// TIA Portal project "Hardware" (V21)

(* hardware
DEVICE "Controller"  S7-1500 station
   slot 0: "Rail_0"  Rack  6ES7 590-1***0-0AA0
   slot 1: "Controller"  CPU 1516-3 PN/DP  6ES7 516-3AN02-0AB0  V2.9
      slot 3: "CPU display_1"  6ES7591-1BA00-0AA0
      slot 32768: "PROFINET interface_1"  X1
         slot 32769: "Port_1"  X1 P1
         slot 32770: "Port_2"  X1 P2
      slot 33024: "PROFINET interface_2"  X2
         slot 33025: "Port_1"  X2 P1
      slot 33280: "DP interface_1"  X3
      slot 34817: "Virtual CP interface port_1"  Virtual CP interface port  Virtual CP interface port
   slot 2: "DI_Main"  DI 32x24VDC HF  6ES7 521-1BL00-0AB0  V2.2
   slot 3: "DQ_Main"  DQ 32x24VDC/0.5A HF  6ES7 522-1BL01-0AB0  V1.1
   slot 4: "AI_Main"  AI 8xU/I/RTD/TC ST  6ES7 531-7KF00-0AB0  V2.2
   slot 5: "AQ_Main"  AQ 4xU/I ST  6ES7 532-5HD00-0AB0  V2.2
DEVICE "Remote_PN_1"  ET 200SP-Station
   slot 0: "Rack_0"  Rack  6ES5 710-8MAx1
   slot 0: "Remote_PN_1"  IM 155-6 PN ST  6ES7 155-6AU01-0BN0  V4.2
   slot 1: "Inputs_1"  DI 8x24VDC ST  6ES7 131-6BF01-0BA0  V0.0
      slot 1: "Inputs_1"  DI 8x24VDC ST
   slot 2: "Outputs_1"  DQ 8x24VDC/0.5A ST  6ES7 132-6BF01-0BA0  V0.0
      slot 1: "Outputs_1"  DQ 8x24VDC/0.5A ST
   slot 3: "Analog_1"  AI 4xI 2-,4-wire ST  6ES7 134-6GD01-0BA1  V2.0
      slot 1: "Analog_1"  AI 4xI 2-,4-wire ST
   slot 127: "BA 2xRJ45"  BA 2xRJ45  6ES7 193-6AR00-0AA0  V0.0
      slot 1: "Port_1"  X1 P1R  6ES7 193-6AR00-0AA0  V0.0
      slot 2: "Port_2"  X1 P2R  6ES7 193-6AR00-0AA0  V0.0
DEVICE "Remote_PN_2"  ET 200SP-Station
   slot 0: "Rack_0"  Rack  6ES5 710-8MAx1
   slot 0: "Remote_PN_2"  IM 155-6 PN ST  6ES7 155-6AU01-0BN0  V4.2
   slot 1: "Inputs_2"  DI 8x24VDC ST  6ES7 131-6BF01-0BA0  V0.0
      slot 1: "Inputs_2"  DI 8x24VDC ST
   slot 127: "BA 2xRJ45"  BA 2xRJ45  6ES7 193-6AR00-0AA0  V0.0
      slot 1: "Port_1"  X1 P1R  6ES7 193-6AR00-0AA0  V0.0
      slot 2: "Port_2"  X1 P2R  6ES7 193-6AR00-0AA0  V0.0
DEVICE "Remote_DP"  ET 200SP-Station
   slot 0: "Rack_0"  Rack  6ES5 710-8MAx1
   slot 0: "Remote_DP"  IM 155-6 DP HF  6ES7 155-6BU01-0CN0  V4.2
   slot 1: "Inputs_DP"  DI 8x24VDC ST  6ES7 131-6BF01-0BA0  V0.0
      slot 1: "Inputs_DP"  DI 8x24VDC ST
   slot 2: "Outputs_DP"  DQ 8x24VDC/0.5A ST  6ES7 132-6BF01-0BA0  V0.0
      slot 1: "Outputs_DP"  DQ 8x24VDC/0.5A ST
DEVICE "Partner"  S7-1500 station
   slot 0: "Rail_0"  Rack  6ES7 590-1***0-0AA0
   slot 1: "Partner"  CPU 1511-1 PN  6ES7 511-1AK02-0AB0  V2.9
      slot 3: "CPU display_1"  6ES7591-1AA00-0AA0
      slot 32768: "PROFINET interface_1"  X1
         slot 32769: "Port_1"  X1 P1
         slot 32770: "Port_2"  X1 P2
      slot 34817: "Virtual CP interface port_1"  Virtual CP interface port  Virtual CP interface port
DEVICE "Partner_IO"  ET 200SP-Station
   slot 0: "Rack_0"  Rack  6ES5 710-8MAx1
   slot 0: "Partner_IO"  IM 155-6 PN ST  6ES7 155-6AU01-0BN0  V4.2
   slot 1: "Outputs_P"  DQ 8x24VDC/0.5A ST  6ES7 132-6BF01-0BA0  V0.0
      slot 1: "Outputs_P"  DQ 8x24VDC/0.5A ST
   slot 127: "BA 2xRJ45"  BA 2xRJ45  6ES7 193-6AR00-0AA0  V0.0
      slot 1: "Port_1"  X1 P1R  6ES7 193-6AR00-0AA0  V0.0
      slot 2: "Port_2"  X1 P2R  6ES7 193-6AR00-0AA0  V0.0
DEVICE "Spare_PN"  ET 200SP-Station
   slot 0: "Rack_0"  Rack  6ES5 710-8MAx1
   slot 0: "Spare_PN"  IM 155-6 PN ST  6ES7 155-6AU01-0BN0  V4.2
   slot 1: "Inputs_S"  DI 8x24VDC ST  6ES7 131-6BF01-0BA0  V0.0
      slot 1: "Inputs_S"  DI 8x24VDC ST
   slot 127: "BA 2xRJ45"  BA 2xRJ45  6ES7 193-6AR00-0AA0  V0.0
      slot 1: "Port_1"  X1 P1R  6ES7 193-6AR00-0AA0  V0.0
      slot 2: "Port_2"  X1 P2R  6ES7 193-6AR00-0AA0  V0.0
*)

// ===== PLC "Controller"  CPU 1516-3 PN/DP =====

VAR_GLOBAL   // PLC tag table "IO"
   "Start_Line" AT %I10.0 : Bool;   // First input of DI_Main
   "Lamp_Line" AT %Q0.0 : Bool;   // First output of DQ_Main
END_VAR

ORGANIZATION_BLOCK "Main"   // OB1, SCL, ProgramCycle
TITLE = "Main Program Sweep (Cycle)"
{ S7_Optimized_Access := 'TRUE' }
VERSION : 0.1
   VAR_INPUT
      Initial_Call : Bool;   // Initial call of this OB
      Remanence : Bool;   // =True, if remanent data are available
   END_VAR
BEGIN

    "Lamp_Line" := "Start_Line";
END_ORGANIZATION_BLOCK

// ===== PLC "Partner"  CPU 1511-1 PN =====

VAR_GLOBAL   // PLC tag table "IO"
   "Start_Partner" AT %I0.0 : Bool;   // An input of the partner
   "Lamp_Partner" AT %Q0.0 : Bool;   // First output of Outputs_P
END_VAR

ORGANIZATION_BLOCK "Main"   // OB1, SCL, ProgramCycle
TITLE = "Main Program Sweep (Cycle)"
{ S7_Optimized_Access := 'TRUE' }
VERSION : 0.1
   VAR_INPUT
      Initial_Call : Bool;   // Initial call of this OB
      Remanence : Bool;   // =True, if remanent data are available
   END_VAR
BEGIN

    "Lamp_Partner" := "Start_Partner";
END_ORGANIZATION_BLOCK